TYPE ST_WorkshopInputs :
STRUCT
    bButton : BOOL;
END_STRUCT
END_TYPE

(* stored: Version 1.1.0.1
   DUT ST_WorkshopInputs: Id {f6ac747e-e3af-4d6a-92d3-a2015627d47e} *)
